// TIA Portal V21 export
// export: Created 2026-11-10T23:32:24.6787448Z, ExportSetting WithDefaults, DisplayName Totally Integrated Automation Portal, DisplayVersion V21 Update 3, DisplayName STEP 7 Professional, DisplayVersion V21 Update 3, DisplayName STEP 7 Safety, DisplayVersion V21, DisplayName Tech WebApplication, DisplayVersion V21, DisplayName WinCC Basic/Comfort/Advanced, DisplayVersion V21 Update 3, DisplayName WinCC Unified, DisplayVersion V21 Update 3
DATA_BLOCK "CamTrack_1"   // DB13, Motion_DB
// stored: AutoNumber true, DBAccessibleFromOPCUA true, DBAccessibleFromWebserver true, InstanceOfName TO_CamTrack, OfSystemLibElement TO_CamTrack, OfSystemLibVersion 8.0
TO_CamTrack   // technology object, version 8.0
// stored: Connection Interface OutputCam
   // // inherited from TO_Object
   // VAR
   //    Parameter { S7_SetPoint := 'True'} : TO_CamTrack_Struct_Parameter;
   //    Interface { S7_SetPoint := 'True'} : TO_CamTrack_Struct_Interface;
   //    Status { ExternalWritable := 'False'} : DInt;
   //    TrackOutput { ExternalWritable := 'False'} : Bool;
   //    SingleCamState { ExternalWritable := 'False'} : DWord;
   //    TrackPosition { ExternalWritable := 'False'} : LReal;
   //    MatchPosition { ExternalWritable := 'False'} : LReal;
   //    Units { ExternalWritable := 'False'; S7_SetPoint := 'True'} : TO_CamTrack_Struct_Units;
   //    StatusWord { ExternalWritable := 'False'} : DWord;
   //    ErrorWord { ExternalWritable := 'False'} : DWord;
   //    ErrorDetail { ExternalWritable := 'False'; S7_SetPoint := 'True'} : TO_Struct_ErrorDetail;
   //    WarningWord { ExternalWritable := 'False'} : DWord;
   // END_VAR
BEGIN
   Parameter.CamTrackLength := 1000.0;
   Parameter.Cam[1..32].Duration := 1.0;
END_DATA_BLOCK
